FUNCTION_BLOCK MissingDestination
  (* Standard: 61499-1; Description: Copyright (c) 2026 Martin Erich Jobst This program and the accompanying materials are made available under the terms of the Eclipse Public License 2.0 which is available at https://www.eclipse.org/legal/epl-2.0/ SPDX-License-Identifier: EPL-2.0 *)
  (* Version 1.0, 2026-11-18, Martin Jobst *)
  PACKAGE lib::Connection;
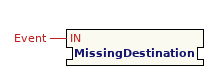
  EVENT_INPUT
    IN;
  END_EVENT
  EVENT_CONNECTIONS
    IN TO Missing.REQ;
  END_CONNECTIONS
END_FUNCTION_BLOCK
